Fanuc KAREL source: kd00043.KL

-- PROVISIONAL review KL for V770-1; original PC SHA256 808ef10d9aca8d580608f1c23d37965cc6d6c472f64a5c8ea62d6e5e2737d24a
-- Incomplete behavior may be omitted. Consult companion uncertainty JSON. Do not deploy.
PROGRAM KD00043
%NOLOCKGROUP
VAR
  I : INTEGER
  J : INTEGER
  B : BOOLEAN
  R : REAL
  S : STRING[80]
-- UNRESOLVED_DECL C type=000014
BEGIN
  -- UNRESOLVED_PC offsets 5-12; opcodes 9D,23
  -- UNRESOLVED_PC offsets 17-21; opcodes 7F
END KD00043
